(* IEC 61131-3 sources: llm-plc-st-eval/data/processed_v2/gpt-4o/B5/zero_shot, 3 files *)

(* ---- ejec_1.st ---- *)
FUNCTION_BLOCK FB_Ventilador
VAR
    // Variable de entrada: estado del quemador
    quemadorOn : BOOL;

    // Variable de salida: estado del ventilador
    ventilador : BOOL;

    // Temporizador para controlar el tiempo de funcionamiento adicional del ventilador
    timer : TON;

    // Variable interna para almacenar el estado previo del quemador
    quemadorPrev : BOOL;
END_VAR

// Inicialización del temporizador
timer(IN := FALSE, PT := T#30S);

// Lógica del ventilador
IF quemadorOn THEN
    // Si el quemador está encendido, el ventilador debe estar encendido
    ventilador := TRUE;
    // Reiniciar el temporizador si el quemador está encendido
    timer(IN := FALSE);
ELSE
    // Si el quemador se apaga, iniciar el temporizador
    IF NOT quemadorPrev THEN
        timer(IN := TRUE);
    END_IF;

    // El ventilador sigue encendido mientras el temporizador está activo
    ventilador := timer.Q;
END_IF;

// Actualizar el estado previo del quemador
quemadorPrev := quemadorOn;
END_FUNCTION_BLOCK

(* ---- ejec_2.st ---- *)
FUNCTION_BLOCK FB_Ventilador
VAR
    // Variable de entrada: indica si el quemador está encendido
    quemadorOn : BOOL;

    // Variable de salida: controla el estado del ventilador
    ventilador : BOOL;

    // Temporizador para controlar el tiempo adicional de funcionamiento del ventilador
    timer : TON;

    // Variable interna para almacenar el estado anterior del quemador
    quemadorPrev : BOOL;
END_VAR

// Inicialización del temporizador
timer(IN := FALSE, PT := T#30S);

// Lógica de control del ventilador
IF quemadorOn THEN
    // Si el quemador está encendido, el ventilador debe estar encendido
    ventilador := TRUE;
    // Reiniciar el temporizador si el quemador está encendido
    timer(IN := FALSE);
ELSE
    // Si el quemador se apaga, iniciar el temporizador
    IF NOT quemadorPrev THEN
        timer(IN := TRUE);
    END_IF;

    // El ventilador sigue encendido mientras el temporizador no haya alcanzado el tiempo preestablecido
    ventilador := NOT timer.Q;
END_IF;

// Actualizar el estado anterior del quemador
quemadorPrev := quemadorOn;
END_FUNCTION_BLOCK

(* ---- ejec_3.st ---- *)
FUNCTION_BLOCK FB_Ventilador
VAR
    // Variable de entrada
    quemadorOn : BOOL; // Estado del quemador: TRUE si está encendido, FALSE si está apagado

    // Variable de salida
    ventilador : BOOL; // Estado del ventilador: TRUE si está encendido, FALSE si está apagado

    // Variables internas
    timer : TON; // Temporizador para controlar el tiempo adicional de funcionamiento del ventilador
END_VAR

// Inicialización del temporizador
timer(IN := NOT quemadorOn, PT := T#30S);

// Lógica de control del ventilador
IF quemadorOn THEN
    ventilador := TRUE; // El ventilador está encendido mientras el quemador está encendido
ELSE
    timer(IN := TRUE); // Iniciar el temporizador cuando el quemador se apaga
    ventilador := timer.Q; // El ventilador sigue encendido mientras el temporizador está activo
END_IF;
